Fanuc KAREL source: KC00006.KL

PROGRAM KC00006
%NOLOCKGROUP
%ENVIRONMENT PBCORE
VAR
  I: INTEGER
  J: INTEGER
  K: INTEGER
  R: REAL
  B: BOOLEAN
  S: STRING[80]
  T: STRING[80]
  P: PATH
  Q: PATH
  AI: ARRAY[8] OF INTEGER
  AB: ARRAY[244] OF BYTE
BEGIN
  APPEND_NODE(P,I)
END KC00006
